// TIA Portal V20 export
Screen "Shapes"  NonexNone, Number=50
  ScreenLayer 
    Rectangle "Rectangle_2" at 624,622 size 254x30
    Line "Line_1" at 174,93 size 480x5
    GraphicView "Graphic view_2" at 27,352 size 140x110  Picture=Graphic_5
